FUNCTION_BLOCK wtch_trend (* Composite Function Block Type *)
  (* Standard: 61499-2 *)
  (* Version 0.0, 12/30/2019, prana, nxtControl GmbH, template *)
  PACKAGE Main;
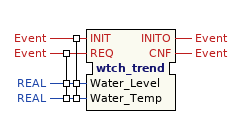
  EVENT_INPUT
    INIT WITH Water_Level, Water_Temp; (* Initialization Request *)
    REQ WITH Water_Level, Water_Temp; (* Normal Execution Request *)
  END_EVENT
  EVENT_OUTPUT
    INITO; (* Initialization Confirm *)
    CNF; (* Execution Confirmation *)
  END_EVENT
  VAR_INPUT
    Water_Level : REAL; (* Input event qualifier *)
    Water_Temp : REAL;
  END_VAR
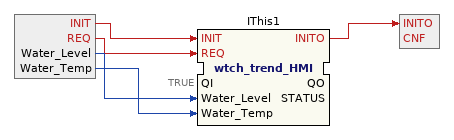
  FBS
    IThis1 : wtch_trend_HMI(QI := TRUE);
  END_FBS
  EVENT_CONNECTIONS
    INIT TO IThis1.INIT;
    REQ TO IThis1.REQ;
    IThis1.INITO TO INITO;
  END_CONNECTIONS
  DATA_CONNECTIONS
    Water_Level TO IThis1.Water_Level;
    Water_Temp TO IThis1.Water_Temp;
  END_CONNECTIONS
END_FUNCTION_BLOCK
